// TIA Portal V21 export
// export: Created 2026-11-10T19:16:51.5147976Z, ExportSetting WithDefaults, DisplayName Totally Integrated Automation Portal, DisplayVersion V21 Update 3, DisplayName STEP 7 Professional, DisplayVersion V21 Update 3, DisplayName STEP 7 Safety, DisplayVersion V21, DisplayName Tech WebApplication, DisplayVersion V21, DisplayName WinCC Basic/Comfort/Advanced, DisplayVersion V21 Update 3, DisplayName WinCC Unified, DisplayVersion V21 Update 3
DATA_BLOCK "FB_Top_DB"   // DB11
VERSION : 0.1
// stored: AutoNumber true, DBAccessibleFromOPCUA true, DBAccessibleFromWebserver true, InstanceOfName FB_Top, InstanceOfType FB
"FB_Top"
   // VAR
   //    "m" { S7_SetPoint := 'True'} : "FB_Multi";
   //    ms { S7_SetPoint := 'True'} : Array[0..1] of "FB_Multi";
   //    x : Real;
   // END_VAR
BEGIN
   "m".sub.stInt := 55;
   ms[0].data.txt := 'deep';
   ms[1].cnt := 9;
END_DATA_BLOCK
